(* IEC 61131-3 sources: s22-soft-shell/st_interpret/tests/test_inputs/st_subset_9_funcs, 2 files *)

(* ---- SimpleAddFunction.st ---- *)
FUNCTION SimpleAddFunction : INT //INT is the return parameter data type
VAR_INPUT
  Input1 :	INT; //Input parameter 1 to the function
  Input2 :	INT; //Input parameter 2 to the function
END_VAR

VAR
  Sum :	INT; //Local variable for temporary calculation
END_VAR

  Sum:= Input1 + Input2; //Total sum

  SimpleAddFunction:= Sum; //Set the return parameter

END_FUNCTION

(* ---- ValueAverageFunction.st ---- *)
FUNCTION ValueAverageFunction : REAL //REAL is the return parameter data type
VAR_INPUT
  Value1 :	REAL; //Input parameter 1 to the function
  Value2 :	REAL; //Input parameter 2 to the function
END_VAR

VAR
  Sum :	REAL; //Local variable for temporary calculation
END_VAR

  Sum:= Value1 + Value2; //Total sum
  Sum:= Sum/2; //Average

  ValueAverageFunction:= Sum; //Set the return parameter

END_FUNCTION
